RoboDK station: minimal.rdk

Station MinStation (saved by RoboDK 6.0.7). Poses are relative to the parent item; angles as X-Y-Z fixed-axis rotations.
  - frame FrameA at (100, 200, 300) mm, rotated rx 0 ry 0 rz 90 deg
    - target TargetB (Cartesian target) at (10, 20, 30) mm; joints []
